(*
	Handles each ended span as soon as the provider hands it over: enrich, then export.
	export clones the span and offers the clone to the exporter as a batch of one. The span is
	dropped when the exporter is busy or the clone fails, and nothing is kept between calls.
	Pass 0 as the exporter to drop every span, or override export to send spans somewhere
	else. Use FB_SpanExporter_Console to write spans to the ADS log.
*)
FUNCTION_BLOCK FB_SpanProcessor_Simple EXTENDS FB_SpanProcessor_Base
VAR
	_spans: FB_SpanQueue(maxCount:=1);
	_exporter: REFERENCE TO FB_SpanExporter_Base;
END_VAR

// no-op; override to change or add to the span before it is exported
METHOD enrich
VAR_IN_OUT
	span: FB_Span;
END_VAR
END_METHOD

(* Sends one ended span on. The span is borrowed for the duration of the call, so the
   exporter is given a clone, which it owns once it accepts it. *)
METHOD export
VAR_INPUT
	span: REFERENCE TO FB_Span;
END_VAR
VAR
	_pClone: POINTER TO FB_Span;
	_cloneFailureReason: E_SpanCloneFailureReason;
	_queueFailureReason: E_SpanQueueFailureReason;
	_exportFailureReason: E_SpanExporterFailureReason;
END_VAR
IF NOT __ISVALIDREF(THIS^._exporter) OR_ELSE THIS^._exporter.isBusy() THEN
	RETURN;
END_IF

IF span.cloneTo(pDest:=_pClone, failureReason=>_cloneFailureReason)
	AND_THEN THIS^._spans.push(pValue:=_pClone, failureReason=>_queueFailureReason) THEN
	THIS^._exporter.export(spans:=THIS^._spans, count:=1, failureReason=>_exportFailureReason);
END_IF

// whatever the exporter did not accept is dropped
THIS^._spans.free();
IF _pClone <> 0 THEN _pClone^.delete(pSelf:=_pClone); END_IF
END_METHOD

METHOD FB_Exit : BOOL
VAR_INPUT
	bInCopyCode: BOOL;  // TRUE: the exit method is called in order to leave the instance which will be copied afterwards (online change).
END_VAR
IF NOT bInCopyCode THEN
	THIS^.free();
END_IF
END_METHOD

// the simple processor keeps nothing between calls; this releases a span left by a failed hand-off
METHOD free
THIS^._spans.free();
END_METHOD

METHOD onEnd
VAR_INPUT
	span: REFERENCE TO FB_Span;
END_VAR
IF NOT __ISVALIDREF(span) THEN
	RETURN;
END_IF

THIS^.enrich(span);
THIS^.export(span);
END_METHOD

// advances the exporter's delivery once per provider tick
METHOD tick
VAR
	_exportFailureReason: E_SpanExporterFailureReason;
END_VAR
IF __ISVALIDREF(THIS^._exporter) THEN
	THIS^._exporter.tick(failureReason=>_exportFailureReason);
END_IF
END_METHOD

METHOD FB_Init : BOOL
VAR_INPUT
	bInitRetains: BOOL;  // TRUE: the retain variables are initialized (reset warm / reset cold)
	bInCopyCode: BOOL;  // TRUE: the instance will be copied to the copy code afterward (online change)
	exporter: REFERENCE TO FB_SpanExporter_Base;  // borrowed and must outlive the processor; 0 drops every span
END_VAR
IF __ISVALIDREF(exporter) THEN
	THIS^._exporter REF= exporter;
ELSE
	THIS^._exporter REF= 0;
END_IF
END_METHOD

END_FUNCTION_BLOCK

(* stored: Version 1.1.0.1
   POU FB_SpanProcessor_Simple: Id {60eb4cc9-96f9-4fec-956a-893d74d004a7}, SpecialFunc None
   Method enrich: Id {c86369c3-3b2f-4cff-9cae-ac60096fe190}
   Method export: Id {e23aeb4f-0578-4d80-920b-0707ff036a41}
   Method FB_Exit: Id {aa794779-2300-4745-90d9-e47ab6a0c9cd}
   Method free: Id {4afad73c-67d9-4058-80c6-cd8d4b6ca5a6}
   Method onEnd: Id {33e9352a-8eea-463d-a646-7a407c79cc74}
   Method tick: Id {ff0bbd46-b17e-4a44-9a5a-c4e4e7871d87}
   Method FB_Init: Id {63177fde-2c04-4e1b-adf4-7d0c9d5c04b4} *)
